// TIA Portal V21 export
TextList "TL_Mode"  ListRange=Decimal
  TextListEntry   Text="-"
  TextListEntry   From=1, To=1, Text="AUTOMATSKI"
  TextListEntry   From=2, To=2, Text="POLUAUTOMATSKI"
  TextListEntry   From=3, To=3, Text="RUČNO"
